Fanuc KAREL source: KO00105.KL

PROGRAM KO00105
%NOLOCKGROUP
VAR
  A: REAL
  B: INTEGER
  OUT: INTEGER
BEGIN
  A = 1
  B = 2
  OUT = ATAN2(A, B)
END KO00105
